FUNCTION_BLOCK AQ_Q_TO_BYTE (* Composite FB for convert AQ to BYTE (QUARTER, 2 Bit) *)
  (* Standard: 61499-2; Description: Copyright (c) 2026 HR Agrartechnik GmbH This program and the accompanying materials are made available under the terms of the Eclipse Public License 2.0 which is available at https://www.eclipse.org/legal/epl-2.0/ SPDX-License-Identifier: EPL-2.0 *)
  (* Version 1.0, 2026-11-13, Franz Höpfinger, HR Agrartechnik GmbH, Initial Version - Luecke geschlossen (analog zu AB_B_TO_BYTE) *)
  PACKAGE adapter::conversion::unidirectional;
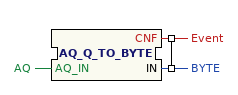
  EVENT_OUTPUT
    CNF WITH IN; (* Confirmation from Adapter *)
  END_EVENT
  VAR_OUTPUT
    IN : BYTE; (* Input data from Adapter *)
  END_VAR
  SOCKETS
    AQ_IN : adapter::types::unidirectional::AQ; (* Adapter Input *)
  END_SOCKETS
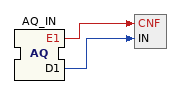
  EVENT_CONNECTIONS
    AQ_IN.E1 TO CNF;
  END_CONNECTIONS
  DATA_CONNECTIONS
    AQ_IN.D1 TO IN;
  END_CONNECTIONS
END_FUNCTION_BLOCK
